Fanuc KAREL source: KA00146.KL

PROGRAM KA00146
%NOLOCKGROUP
VAR
  SRC: ARRAY[4] OF INTEGER
  DST: ARRAY[4] OF REAL
BEGIN
  DST = SRC
END KA00146
